INTERFACE I_MoverEnableAlgorithm EXTENDS i_Task


METHOD Abort : HRESULT
VAR_INPUT
END_VAR
END_METHOD

METHOD Enable : HRESULT
VAR_INPUT
END_VAR
END_METHOD

METHOD Reset : HRESULT
VAR_INPUT
END_VAR
END_METHOD

METHOD SetComponents : BOOL
VAR_INPUT
	MoverArray : ARRAY[0..TcIoXtsEnvironmentParameterList.MaxXtsMoversPerXpu] OF I_XtsMover;
	CAGroup : I_CollisionGroup;
	MoverCount : UDINT;
END_VAR
END_METHOD

END_INTERFACE

(* stored: Version 1.1.0.1
   Itf I_MoverEnableAlgorithm: Id {fc5ea72b-09f8-4cbb-94b5-463ddba58f35}
   Method Abort: Id {b0bc9a74-deef-4234-b8f9-c8c9d46ad2c9}
   Method Enable: Id {1180b379-2462-48af-a710-0e37d3d9156e}
   Method Reset: Id {0f25d9f6-907a-4ed5-8a8f-75e5bc9f2b4b}
   Method SetComponents: Id {8f66a473-b73c-4779-bff7-f5bae82d2f36} *)
